(* IEC 61131-3 sources: st-fmt/tests/fixtures/types, 2 files *)

(* ---- type_block.expected.st ---- *)
TYPE
Point : STRUCT
    x     : REAL;
    y     : REAL;
    label : STRING[32] := '';
END_STRUCT

Overlay : UNION
    bits  : DWORD;
    value : REAL;
END_UNION

Meters : INT (0..100);
Alias : ARRAY [0..9] OF INT;
Color : (Red, Green, Blue);
State : (
    Idle    := 0,
    Running := 10,
    Faulted := 20,
);
Counter : UDINT := 0;
END_TYPE

(* ---- type_block.st ---- *)
type
Point : struct
x : real;
y : real;
label : STRING[32] := '';
end_struct

Overlay : union
bits : dword;
value : real;
end_union

Meters : INT (0..100);
Alias : ARRAY [0..9] OF int;
Color : (Red, Green, Blue);
State : (Idle := 0, Running := 10, Faulted := 20);
Counter : udint := 0;
end_type
